Fanuc KAREL source: kf00098.KL

-- PROVISIONAL review KL for V1013-1; original PC SHA256 6cb9920c8af5ba8f0446998c487e4732e44b8600fcc38f100c96dae94577bedb
-- Incomplete behavior may be omitted. Consult companion uncertainty JSON. Do not deploy.
PROGRAM KF00098
%NOLOCKGROUP
BEGIN
  -- UNRESOLVED_PC offsets 5-16; opcodes 2E,23
  -- UNRESOLVED_PC offsets 21-32; opcodes 2E,23
  -- UNRESOLVED_PC offsets 37-55; opcodes 27,27,9D,22,22,31
  -- UNRESOLVED_PC offsets 60-64; opcodes 7F
END KF00098
